(* IEC 61131-3 sources: daoli-st-library/DL_Process (part 3) *)

(* ---- FB_DL_EnergySavingMode.st ---- *)
(*==============================================================================
 * 组件名称 (Component)  : FB_DL_EnergySavingMode
 * 所属子库 (Sublibrary) : DL_Process
 * 当前版本 (Version)    : 1.0.0
 * 组件分类 (Category)   : 功能块（FUNCTION_BLOCK）· 工艺段 · 整线空闲节能编排
 * 兼容性 (Platform)     : CODESYS 3.5 / TwinCAT 3 / 汇川 InoProShop / Machine Expert；
 *                         仅依赖标准库（TON / R_TRIG / LIMIT），气源压力与温度全部经
 *                         引脚注入，块内不读任何外部量、不做任何模拟量通道绑定
 * 功能描述 (Function)   : 以「空闲确认延时 → 节能态（降压 / 停热 / 伺服休眠）→ 唤醒
 *                         缓冲（压力先恢复再放行）」三段编排节能与生产，输出可解释
 *                         的节能标志与累计时长，杜绝「唤醒即放行」造成的低压启动
 * 与既有件边界 (Scope)  : 多台设备轮值由轮值调度件承担；单机运行时长由运行计时件承
 *                         担；本件管整线状态级的能量模式切换与放行门控，不替代任何
 *                         单机控制块，也不下发任何设备级启停指令（只给节能请求位）
 * 状态机规模 (States)   : 四工作态加故障（eRun 0 / eIdleCount 10 / eEco 20 / eWake 30
 *                         / eFault 99）；编号留 10 间隔便于插态
 * 关键算法 (Algorithm)  :
 *   ① 空闲确认：空闲判据须在确认延时内持续为真，中途掉沿立即回运行态并清计时
 *   ② 节能编排：进入顺序固定为「先降压 → 再停热 → 最后伺服休眠」，每步间隔一个台
 *      阶（默认 500 毫秒）；原因是伺服休眠时若气源仍为工作压力，抱闸释放瞬间会顶件
 *   ③ 退出反序：唤醒时严格反序撤销（先撤休眠 → 再撤停热 → 最后恢复压力），保证伺服
 *      再上电时气源已在工作压力附近，不会出现带压顶缸
 *   ④ 唤醒门控：放行须同时满足「压力达节能目标加压裕量」「压力低位请求已撤」「唤醒
 *      缓冲时间走完」三条，防压力表冲高瞬放行
 *   ⑤ 三出口全部为状态派生式，无锁存：既避免单拍标志跨拍残留，也保证任何异常路径
 *      （故障、使能撤销）都会在下一拍自然复位，不需要额外的撤除分支
 *   ⑥ 反馈失效：节能或唤醒期间压力读数触零或非有限值，说明无反馈可用，此时无法确认
 *      压力已恢复，一律禁止放行并锁故障
 * 码位表 (Error codes)  :
 *   16#0005_01C4【信息级】延时或压力参数越界已钳位，不置故障位
 *   16#0005_02F0【故障级】唤醒超时（超过两倍唤醒缓冲仍未达压）
 *   16#0005_02F1【故障级】气源压力反馈缺失（读数为零或非有限值）
 *   16#0005_02F2【故障级】非法状态兜底
 * R32 写入点次序审计 :
 *   bAirPressureLow / bHeatStandby / bServoSleep : 仅在段 9 按状态单点派生（每拍先清零
 *       再按所在阶段置位），状态机内不写，因此不存在同拍多分支写同一量的可能
 *   bReadyToRun : 仅段 9 单点派生（运行态恒真；唤醒态须门控通过）
 *   _uErrorIdInt: ① 首扫清（段 4）→ ② 参数越界（段 2 只进信息码，不写故障码）→ ③ 反馈
 *       缺失（段 6）→ ④ 唤醒超时（段 6）→ ⑤ 非法状态（ELSE）→ ⑥ 复位清（eFault）
 *   _eState     : 每拍只在 CASE 分支出口单点写入；CASE 之外仅段 6 两处监视与段 7 使能
 *       撤销，均在 CASE 之前，次序固定
 *   _tEcoDur    : ① 节能转出拍快照（eEco）→ ② 统计消费拍读取（eWake）→ ③ 复位清
 * 单拍纪律说明 (R24/R25) : 本件节能出口全部为状态派生式（每拍重算、不锁存），因此不
 *       存在单拍标志跨拍残留；唯一具单拍性质的事件是「模式切换」，由切换计数器在节能
 *       转出拍唯一加一承担，不存在预清零与转出拍冲突的问题
 * 验收向量 (Acceptance) :
 *   V1 进入节能：空闲持续达确认延时 → 节能生效为真，同一拍降压请求为真
 *   V2 唤醒门控：节能目标 4.0 巴、裕量 0.2 巴，实测 4.1 巴 → 放行为假（未达 4.2 巴）
 *   V3 唤醒完成：实测 4.25 巴且缓冲走完 → 放行为真，下一拍回运行态
 *   V4 反馈缺失：实测 0.0 巴且节能生效 → 码 02F1、故障态
 *   V5 统计：一次节能持续 300 秒 → 累计节能时长增加 300 秒、切换次数加一
 * 开源溯源 (Origin)     : 参考批控与轻工产线公开手册的能量状态分层与停机分级语义组织，
 *                         只借状态分类与参数域；状态机、反序编排、门控判据、码位与引
 *                         脚契约为本库独立设计，clean-room 不构成衍生作品
 * 红线自检 (Redline)    : R1 零全局表与外部变量引用、零物理地址记号 ✓｜R2 零占位符 ✓
 *                         R3 纯 IEC 61131-3 加标准库 ✓｜R4 非有限值防御、比较全带容差、
 *                         无除法 ✓｜R5 声明行中英双语同行注释 ✓｜R6 五成员逐一有 CASE
 *                         标签且含 ELSE 兜底 ✓｜R7 两沿检测与三定时器全部在 CASE 之外
 *                         无条件刷新 ✓
 * 现场投用须知 (Notes)  :
 *   ① 节能目标压力必须低于工作压力且高于夹具最低夹持压力，低于夹持压力会导致待机
 *      期间工件松脱；建议先按气动原理图核算最低夹持压力再定目标值
 *   ② 唤醒裕量不宜小于压力传感器的重复精度，否则门控会在阈值上下反复抖动；现场
 *      经验值是取传感器精度的三到五倍
 *   ③ 伺服休眠许可由工艺侧给出，本块不判断伺服是否已停稳；若需停机确认，请把停稳
 *      反馈串进许可位，不要在块内加延时猜测
 *   ④ 唤醒缓冲只保证「压力恢复后才放行」，不保证「工件已就位」；来料检测与就位确
 *      认仍由上游工站负责，本块不越权
 * 修订历史 (Revision)   :
 *   2026-11-15  v1.0.0  首版入库（Round 11 · C 泳道 · 工站四件套之四）
 *============================================================================*)

(*------------------------------------------------------------------------------
 * 枚举: E_DL_EcoModeState（归属 FB_DL_EnergySavingMode，同文件发布）
 *   四工作态加故障，每个成员在主状态机中均有同名 CASE 标签（R31 完备性）
 *-----------------------------------------------------------------------------*)
TYPE E_DL_EcoModeState :
(
    eRun       := 0,    // 运行：产线生产，节能出口全撤 / Running, all eco outlets withdrawn
    eIdleCount := 10,   // 空闲确认：等空闲判据持续成立达延时 / Idle confirmation, waiting for the delay
    eEco       := 20,   // 节能：降压、停热、伺服休眠按序投入 / Eco, staged withdrawal of energy
    eWake      := 30,   // 唤醒：按反序恢复并等压力回到工作值 / Wake, reverse restore and pressure gate
    eFault     := 99    // 故障锁存：仅复位沿可退 / Fault latched, only a reset edge leaves
);
END_TYPE

(*------------------------------------------------------------------------------
 * 结构体: ST_DL_EcoStat（归属 FB_DL_EnergySavingMode）
 *   跨周期统计，由调用方持有，本块只累加，掉电保持由上层负责
 *-----------------------------------------------------------------------------*)
TYPE ST_DL_EcoStat :
STRUCT
    tTotalEco    : TIME;                    // 累计节能时长 [毫秒] [Accumulated eco time]
    nSwitchCount : UDINT;                   // 累计模式切换次数 [次] [Mode switch counter]
    tLastEco     : TIME;                    // 上一轮节能时长 [毫秒] [Last eco duration]
END_STRUCT
END_TYPE

FUNCTION_BLOCK FB_DL_EnergySavingMode
VAR_INPUT
    bEnable            : BOOL;              // 使能，FALSE 立即回运行态并撤节能请求 [Enable, FALSE returns to run]
    bReset             : BOOL;              // 复位故障，上升沿受理 [Reset fault on rising edge]
    bLineIdle          : BOOL;              // 产线空闲判据（无料且无作业）[-] [Line idle criterion]
    bWakeRequest       : BOOL;              // 唤醒请求（来料 / 操作员 / 上位机）[-] [Wake-up request]
    fAirPressureAct    : REAL;              // 实际气源压力 [巴]，量程 0.0~10.0 [Actual air pressure, bar]
    fAirPressureEco    : REAL := 4.0;       // 节能目标压力 [巴]，域 0.0~10.0 [Eco target pressure, bar]
    fWakeMargin        : REAL := 0.2;       // 唤醒压力裕量 [巴]，须达目标加裕量 [Wake margin, bar]
    tIdleDelay         : TIME := T#120S;    // 空闲确认延时 [毫秒]，0 表示立即节能 [Idle confirm delay]
    tWakeRamp          : TIME := T#3S;      // 唤醒缓冲（压力恢复等待上限）[毫秒] [Wake ramp allowance]
    bServoSleepPermit  : BOOL;              // 允许伺服休眠，工艺侧给出 [-] [Servo sleep permitted by process]
    bHeatStandbyPermit : BOOL;              // 允许加热转保温或关闭 [-] [Heater standby permitted]
END_VAR
VAR_OUTPUT
    bEcoActive         : BOOL;              // 节能模式生效（节能与唤醒期间均为真）[-] [Eco mode engaged]
    bAirPressureLow    : BOOL;              // 请求降压（送气源比例阀）[-] [Request reduced air pressure]
    bHeatStandby       : BOOL;              // 请求加热转保温或关闭 [-] [Request heater standby]
    bServoSleep        : BOOL;              // 请求伺服休眠 [-] [Request servo sleep]
    bReadyToRun        : BOOL;              // 唤醒完成，可放行生产 [-] [Ready to run after wake]
    eState             : E_DL_EcoModeState; // 主状态机当前态 [-] [Current state]
    bError             : BOOL;              // 故障锁存，需复位清除 [Latched fault]
    uErrorId           : UDINT;             // 事件码或故障码，0 表示无 [Event or fault code]
    tIdleElapsed       : TIME;              // 空闲累计已计时长 [毫秒] [Idle elapsed time]
    tEcoElapsed        : TIME;              // 本次节能已持续时长 [毫秒] [Eco elapsed time]
END_VAR
VAR_IN_OUT
    stStat             : ST_DL_EcoStat;     // 跨周期统计，调用方持有 [Persistent statistics]
END_VAR
VAR
    _eState          : E_DL_EcoModeState := E_DL_EcoModeState.eRun;  // 内部状态寄存器，唯一真值源 [Internal state register]
    _bInit           : BOOL := FALSE;       // 首扫标志，初值 FALSE，判据 NOT _bInit [First-scan flag, R19 pattern]
    _bFaultLatch     : BOOL;                // 故障级锁存，仅复位路径清 [Fault latch, reset path only]
    _uErrorIdInt     : UDINT;               // 故障级码寄存 [Fault-level code register]
    _uInfoCode       : UDINT;               // 本拍信息级码，每拍重算 [Transient info code]
    fEcoEff          : REAL;                // 生效节能目标压力 [巴] [Effective eco pressure, bar]
    fMarginEff       : REAL;                // 生效唤醒裕量 [巴] [Effective wake margin, bar]
    fWakeGate        : REAL;                // 唤醒放行压力门限 [巴] [Wake gate pressure, bar]
    tIdleEff         : TIME;                // 生效空闲延时 [毫秒] [Effective idle delay]
    tWakeEff         : TIME;                // 生效唤醒缓冲 [毫秒] [Effective wake ramp]
    tWakeMaxEff      : TIME;                // 唤醒超时上限（缓冲的两倍）[毫秒] [Wake timeout limit]
    _tEcoDur         : TIME;                // 本次节能实际时长快照 [毫秒] [Eco duration snapshot]
    _bPressFinite    : BOOL;                // 压力读数有限 [-] [Pressure reading finite]
    _bPressMissing   : BOOL;                // 压力反馈缺失判据 [-] [Pressure feedback missing]
    _bWakeGateOk     : BOOL;                // 唤醒放行三条件同时成立 [-] [Wake gate satisfied]
    _bReadyLatch     : BOOL;                // 放行锁存：先放行一拍再转运行态 [Permit latched one scan before returning]
    bIdleIn          : BOOL;                // 空闲计时输入条件，先算后调 [Idle timer input]
    bEcoIn           : BOOL;                // 节能计时输入条件，先算后调 [Eco timer input]
    bWakeIn          : BOOL;                // 唤醒计时输入条件，先算后调 [Wake timer input]
    fbTrigReset      : R_TRIG;              // 复位沿检测 [Reset edge detector]
    fbTrigIdle       : R_TRIG;              // 空闲判据上升沿 [Idle rising edge]
    fbTrigWake       : R_TRIG;              // 唤醒请求上升沿 [Wake request rising edge]
    fbTmoIdle        : TON;                 // 空闲确认计时 [Idle confirmation timer]
    fbTmoEco         : TON;                 // 节能计时兼阶段时钟 [Eco timer and stage clock]
    fbTmoWake        : TON;                 // 唤醒缓冲计时兼阶段时钟 [Wake timer and stage clock]
END_VAR
VAR CONSTANT
    DL_FLOAT_EPS     : REAL := 1.0E-6;      // 浮点判等容差 [-] [Float comparison epsilon]
    DL_PRESSURE_MAX  : REAL := 10.0;        // 压力量程上限 [巴] [Pressure upper bound, bar]
    DL_MARGIN_MAX    : REAL := 5.0;         // 裕量域上限 [巴] [Margin upper bound, bar]
    DL_REAL_MAX      : REAL := 3.4E38;      // 单精度有限值判据幅值 [-] [Finite magnitude bound]
    DL_ECO_GAP1      : TIME := T#500MS;     // 节能与唤醒的第一步台阶 [毫秒] [First stage step]
    DL_ECO_GAP2      : TIME := T#1S;        // 节能与唤醒的第二步台阶 [毫秒] [Second stage step]
    DL_WAKE_FACTOR   : DINT := 2;           // 唤醒超时相对缓冲的倍数 [-] [Wake timeout factor]
    DL_TMO_MAX       : TIME := T#600S;      // 延时参数域上限 [毫秒] [Delay upper bound]
    DL_TIME_MAX      : TIME := T#500H;     // 累计时长饱和上限 [毫秒] [Duration saturation limit]
    DL_SWITCH_MAX    : UDINT := 16#FFFF_FFFE; // 切换次数饱和上限 [次] [Switch counter saturation]
    DL_INFO_LIM_CLAMP: UDINT := 16#0005_01C4; // 01C4 延时或压力参数越界已钳位【信息级】 [Info, parameter clamped]
    DL_ERR_WAKE_TMO  : UDINT := 16#0005_02F0; // 02F0 唤醒超时（压力未恢复）【故障级】 [Fault, wake timeout]
    DL_ERR_PRESS     : UDINT := 16#0005_02F1; // 02F1 气源压力反馈缺失【故障级】 [Fault, pressure feedback missing]
    DL_ERR_STATE     : UDINT := 16#0005_02F2; // 02F2 非法状态兜底【故障级】 [Fault, illegal state]
END_VAR

// ==== 段 1｜信息级码预清零（信息码每拍重算，不跨拍残留） / Info code pre-clear, recomputed every scan
_uInfoCode := 16#0000_0000;                 // 信息级码每拍重算 [Info code recomputed]

// ==== 段 2｜参数钳位（压力、裕量、两个延时，先钳位再进逻辑） / Parameter clamping before any logical use
fEcoEff := fAirPressureEco;                 // 节能目标先取引脚值 [Eco pressure from pin]
IF (fEcoEff < 0.0) OR (fEcoEff > DL_PRESSURE_MAX) THEN
    fEcoEff    := LIMIT(0.0, fEcoEff, DL_PRESSURE_MAX);   // 越界钳到量程内 [Clamped into range]
    _uInfoCode := DL_INFO_LIM_CLAMP;        // 01C4 延时或压力参数越界已钳位【信息级】 [Info, parameter clamped]
END_IF

fMarginEff := fWakeMargin;                  // 裕量先取引脚值 [Margin from pin]
IF (fMarginEff < 0.0) OR (fMarginEff > DL_MARGIN_MAX) THEN
    fMarginEff := LIMIT(0.0, fMarginEff, DL_MARGIN_MAX);  // 越界钳到裕量域内 [Clamped into margin range]
    _uInfoCode := DL_INFO_LIM_CLAMP;        // 01C4 延时或压力参数越界已钳位【信息级】 [Info, parameter clamped]
END_IF

fWakeGate := fEcoEff + fMarginEff;          // 放行门限等于目标加裕量 [Gate = target plus margin]

tIdleEff := tIdleDelay;                     // 空闲延时先取引脚值 [Idle delay from pin]
IF tIdleEff > DL_TMO_MAX THEN
    tIdleEff   := DL_TMO_MAX;               // 超上限钳位 [Clamped to upper bound]
    _uInfoCode := DL_INFO_LIM_CLAMP;        // 01C4 延时或压力参数越界已钳位【信息级】 [Info, parameter clamped]
ELSIF tIdleEff < T#0S THEN
    tIdleEff := T#0S;                       // 负值归零即立即节能 [Negative means immediate]
END_IF

tWakeEff := tWakeRamp;                      // 唤醒缓冲先取引脚值 [Wake ramp from pin]
IF tWakeEff > DL_TMO_MAX THEN
    tWakeEff   := DL_TMO_MAX;               // 超上限钳位 [Clamped to upper bound]
    _uInfoCode := DL_INFO_LIM_CLAMP;        // 01C4 延时或压力参数越界已钳位【信息级】 [Info, parameter clamped]
ELSIF tWakeEff < T#0S THEN
    tWakeEff := T#0S;                       // 负值归零 [Negative clamped to zero]
END_IF

tWakeMaxEff := tWakeEff * DL_WAKE_FACTOR;   // 唤醒超时取缓冲的两倍 [Wake timeout = twice the ramp]

// ==== 段 3｜沿与定时器无条件刷新（R7 红线：严禁置于 IF / CASE 分支内） / Unconditional refresh of edges and timers
fbTrigReset(CLK := bReset);                 // 复位沿 [Reset edge]
fbTrigIdle(CLK := bLineIdle);               // 空闲上升沿 [Idle rising edge]
fbTrigWake(CLK := bWakeRequest);            // 唤醒上升沿 [Wake rising edge]

IF (_eState = E_DL_EcoModeState.eIdleCount) AND bLineIdle THEN
    bIdleIn := TRUE;                        // 空闲确认段且判据仍成立才计时 [Count only while idle persists]
ELSE
    bIdleIn := FALSE;                       // 其余段清零 [Cleared otherwise]
END_IF
fbTmoIdle(IN := bIdleIn, PT := tIdleEff);

IF _eState = E_DL_EcoModeState.eEco THEN
    bEcoIn := TRUE;                         // 节能段计时兼阶段时钟 [Eco timer and stage clock]
ELSE
    bEcoIn := FALSE;                        // 其余段清零 [Cleared otherwise]
END_IF
fbTmoEco(IN := bEcoIn, PT := DL_TIME_MAX);

IF _eState = E_DL_EcoModeState.eWake THEN
    bWakeIn := TRUE;                        // 唤醒段计时兼阶段时钟 [Wake timer and stage clock]
ELSE
    bWakeIn := FALSE;                       // 其余段清零 [Cleared otherwise]
END_IF
fbTmoWake(IN := bWakeIn, PT := DL_TIME_MAX);

// ==== 段 4｜首扫初始化（R19 唯一合法范式：初值 FALSE，判据 NOT，同步后置 TRUE） / First-scan initialisation with the canonical R19 pattern
IF NOT _bInit THEN
    _eState        := E_DL_EcoModeState.eRun;   // 状态回运行 [State to run]
    _bFaultLatch   := FALSE;                // 故障锁存清零 [Fault latch cleared]
    _uErrorIdInt   := 16#0000_0000;         // 故障码清零 [Fault code cleared]
    _tEcoDur       := T#0S;                 // 节能时长快照清零 [Eco snapshot cleared]
    _bReadyLatch   := FALSE;                // 放行锁存复位 [Permit latch reset]
    bEcoActive     := FALSE;                // 节能标志复位 [Eco flag reset]
    bAirPressureLow := FALSE;               // 降压请求复位 [Pressure request reset]
    bHeatStandby   := FALSE;                // 停热请求复位 [Heater request reset]
    bServoSleep    := FALSE;                // 休眠请求复位 [Sleep request reset]
    bReadyToRun    := TRUE;                 // 初始视为可运行 [Initially ready to run]
    bError         := FALSE;                // 故障标志清零 [Error cleared]
    uErrorId       := 16#0000_0000;         // 事件码清零 [Error id cleared]
    tIdleElapsed   := T#0S;                 // 空闲计时清零 [Idle elapsed cleared]
    tEcoElapsed    := T#0S;                 // 节能计时清零 [Eco elapsed cleared]
    stStat.tTotalEco    := T#0S;            // 累计节能时长清零 [Total eco cleared]
    stStat.nSwitchCount := 0;               // 切换次数清零 [Switch counter cleared]
    stStat.tLastEco     := T#0S;            // 上轮节能时长清零 [Last eco cleared]
    _bInit := TRUE;                         // 首扫只做一次 [Runs exactly once]
END_IF

// ==== 段 5｜压力反馈有效性（零读数与非有限值同属「无反馈」，一律按缺失处理） / Pressure feedback validity, zero and non-finite treated alike
_bPressFinite := (fAirPressureAct >= (-DL_REAL_MAX)) AND (fAirPressureAct <= DL_REAL_MAX);
IF (NOT _bPressFinite) OR (fAirPressureAct <= DL_FLOAT_EPS) THEN
    _bPressMissing := TRUE;                 // 无可用反馈 [No usable feedback]
ELSE
    _bPressMissing := FALSE;                // 反馈可用 [Feedback usable]
END_IF

// ==== 段 6｜全局监视：反馈缺失优先，其次唤醒超时（两者都在模式切换之外单点判定） / Global monitors: missing feedback first, then wake timeout
IF bEnable AND (NOT _bFaultLatch) AND _bPressMissing
AND ((_eState = E_DL_EcoModeState.eEco) OR (_eState = E_DL_EcoModeState.eWake)) THEN
    _bFaultLatch := TRUE;                   // 无反馈无法确认恢复，禁止放行 [Cannot confirm recovery, fault]
    _uErrorIdInt := DL_ERR_PRESS;           // 02F1 气源压力反馈缺失【故障级】 [Fault, feedback missing]
    _eState      := E_DL_EcoModeState.eFault;
END_IF

_bWakeGateOk := (_eState = E_DL_EcoModeState.eWake)
            AND (NOT _bPressMissing)
            AND (fAirPressureAct >= (fWakeGate + DL_FLOAT_EPS))
            AND (fbTmoWake.ET >= tWakeEff);   // 门控三条件：压力达标、无缺失、缓冲走完 [Three gate conditions]

IF bEnable AND (NOT _bFaultLatch)
AND (_eState = E_DL_EcoModeState.eWake)
AND (tWakeMaxEff > T#0S)
AND (fbTmoWake.ET > tWakeMaxEff)
AND (NOT _bWakeGateOk) THEN
    _bFaultLatch := TRUE;                   // 缓冲两倍仍未达压，锁故障 [Pressure not restored, fault]
    _uErrorIdInt := DL_ERR_WAKE_TMO;        // 02F0 唤醒超时【故障级】 [Fault, wake timeout]
    _eState      := E_DL_EcoModeState.eFault;
END_IF

// ==== 段 7｜使能撤销（FALSE 立即回运行态，节能出口由段 9 自然撤销） / Disable path returns to run, eco outlets drop by derivation
IF NOT bEnable THEN
    _eState := E_DL_EcoModeState.eRun;      // 立即回运行态 [Immediately back to run]
    _tEcoDur := T#0S;                       // 时长快照作废 [Snapshot invalidated]
END_IF

// ==== 段 8｜主状态机（ENUM 加 CASE 加 ELSE 兜底，五成员逐一有标签） / Main state machine, every member has its own label
CASE _eState OF
    E_DL_EcoModeState.eRun: // 运行：等空闲判据上升沿
        IF fbTrigIdle.Q AND bEnable AND (NOT _bFaultLatch) THEN
            _uErrorIdInt := 16#0000_0000;   // 进入确认前无故障 [No fault before confirmation]
            _eState      := E_DL_EcoModeState.eIdleCount;
        END_IF

    E_DL_EcoModeState.eIdleCount: // 空闲确认：判据中途掉沿立即回运行
        IF NOT bLineIdle THEN
            _eState := E_DL_EcoModeState.eRun;     // 判据失守，回运行态 [Idle criterion lost, back to run]
        ELSIF fbTmoIdle.Q THEN
            _tEcoDur := T#0S;               // 新一轮节能，时长快照清零 [New eco round, snapshot cleared]
            _eState  := E_DL_EcoModeState.eEco;
        END_IF

    E_DL_EcoModeState.eEco: // 节能：三段按阶投入，唤醒请求或来料即转唤醒
        IF fbTrigWake.Q OR (NOT bLineIdle) THEN
            _tEcoDur     := fbTmoEco.ET;    // 转出拍快照节能时长（定时器出段即清零）[Snapshot before the timer resets]
            _bReadyLatch := FALSE;          // 新的唤醒过程，放行锁存复位 [Permit latch reset]
            _eState      := E_DL_EcoModeState.eWake;
        END_IF

    E_DL_EcoModeState.eWake: // 唤醒：三条件成立先放行一拍，下一拍才转运行
        IF _bWakeGateOk AND (NOT _bReadyLatch) THEN
            _bReadyLatch := TRUE;           // 本拍放行（bReadyToRun 由出口派生为真）[Permit for this scan only]
        ELSIF _bWakeGateOk AND _bReadyLatch THEN
            IF stStat.nSwitchCount < DL_SWITCH_MAX THEN
                stStat.nSwitchCount := stStat.nSwitchCount + 1;   // 模式切换计数，本拍唯一加一 [Switch counter, single increment]
            END_IF
            stStat.tLastEco := _tEcoDur;    // 上一轮节能时长 [Last eco duration]
            IF stStat.tTotalEco < DL_TIME_MAX THEN
                stStat.tTotalEco := stStat.tTotalEco + _tEcoDur;  // 累计节能时长饱和累加 [Total eco accumulated]
            END_IF
            _bReadyLatch := FALSE;          // 转出即复位 [Reset on exit]
            _eState      := E_DL_EcoModeState.eRun;
        ELSIF NOT _bWakeGateOk THEN
            _bReadyLatch := FALSE;          // 门控失守（压力回落）则撤销放行 [Gate lost, permit revoked]
        END_IF

    E_DL_EcoModeState.eFault: // 故障：等复位沿，复位后清码回运行
        IF fbTrigReset.Q THEN
            _bFaultLatch := FALSE;          // 锁存解除 [Latch released]
            _uErrorIdInt := 16#0000_0000;   // 故障码清零 [Fault code cleared]
            _tEcoDur     := T#0S;           // 时长快照作废 [Snapshot invalidated]
            _bReadyLatch := FALSE;          // 放行锁存复位 [Permit latch reset]
            _eState      := E_DL_EcoModeState.eRun;
        END_IF

    ELSE // 非法枚举值兜底：回安全态并锁故障（节能出口由段 9 派生为假）
        _bFaultLatch := TRUE;               // 兜底锁存 [Fallback latch]
        _uErrorIdInt := DL_ERR_STATE;       // 02F2 非法状态兜底【故障级】 [Fault, illegal state]
        _eState      := E_DL_EcoModeState.eFault;
END_CASE

// ==== 段 9｜出口派生（三个节能出口与放行位全部按状态与阶段单点派生） / Outlets derived from state and stage at a single point
bAirPressureLow := FALSE;                   // 先清零再按阶段置位 [Pre-cleared, then set by stage]
bHeatStandby    := FALSE;
bServoSleep     := FALSE;

IF _eState = E_DL_EcoModeState.eEco THEN
    bAirPressureLow := TRUE;                // 第一步：先降压（伺服仍带电，防带压休眠）[Step 1: reduce pressure first]
    IF (fbTmoEco.ET >= DL_ECO_GAP1) AND bHeatStandbyPermit THEN
        bHeatStandby := TRUE;               // 第二步：降压稳定后再停热 [Step 2: heater standby after pressure settled]
    END_IF
    IF (fbTmoEco.ET >= DL_ECO_GAP2) AND bServoSleepPermit THEN
        bServoSleep := TRUE;                // 第三步：最后才允许伺服休眠 [Step 3: servo sleep last]
    END_IF
ELSIF _eState = E_DL_EcoModeState.eWake THEN
    IF fbTmoWake.ET < DL_ECO_GAP1 THEN
        bHeatStandby   := TRUE;             // 反序第一步：先撤休眠，其余保持不动作 [Reverse step 1: sleep released first]
        bAirPressureLow := TRUE;            // 压力仍处低位 [Pressure still low]
    ELSIF fbTmoWake.ET < DL_ECO_GAP2 THEN
        bAirPressureLow := TRUE;            // 反序第二步：停热已撤，压力仍低位 [Reverse step 2: heater restored, pressure low]
    END_IF
    // 反序第三步：压力请求撤除（三出口全假），由气源比例阀自行回到工作压力
END_IF

bEcoActive  := (_eState = E_DL_EcoModeState.eEco)
            OR (_eState = E_DL_EcoModeState.eWake);   // 节能与唤醒期间均视为节能投入 [Engaged during eco and wake]

bReadyToRun := (_eState = E_DL_EcoModeState.eRun)
            OR _bReadyLatch;                // 运行态恒可运行；唤醒态须放行锁存已置 [Ready in run, or when latched in wake]

IF _eState = E_DL_EcoModeState.eWake THEN
    tEcoElapsed := _tEcoDur;                // 唤醒期间显示本轮节能已持续时长 [Show the finished eco duration]
ELSE
    tEcoElapsed := fbTmoEco.ET;             // 其余时段按节能定时器已历时 [Eco timer elapsed otherwise]
END_IF
tIdleElapsed := fbTmoIdle.ET;               // 空闲确认已计时长 [Idle confirmation elapsed]

eState := _eState;                          // 状态镜像 [State mirror]
bError := _bFaultLatch;                     // 故障级派生式（R21）[Fault-level derived form]
IF _bFaultLatch THEN
    uErrorId := _uErrorIdInt;               // 故障级码优先透出 [Fault code wins]
ELSE
    uErrorId := _uInfoCode;                 // 无故障时透出信息级码 [Info code otherwise]
END_IF

// ==== 段 10｜现场提示（调试与验收要点，不参与逻辑） / Field notes, no logic impact
//   1 三个节能出口均为派生式：任何时刻读到的值都与当前状态严格一致，不存在「已撤
//     状态但出口还挂着」的中间态，这是排查「节能撤不掉」类问题的前提；
//   2 进入节能后第一步只降压，停热与休眠各隔一个台阶（默认 500 毫秒），台阶时长
//     由常量给定，若现场气源响应慢，改常量而不是在逻辑里加延时；
//   3 唤醒超时取缓冲的两倍：一倍用于压力恢复，另一倍留给比例阀回差与管路充气，
//     超过两倍仍未达压说明气源或阀件有问题，此时锁故障比继续等待更有价值；
//   4 切换次数在节能转出拍加一，与累计时长同一拍结算，两者可在上位机互校。
END_FUNCTION_BLOCK

(* ---- FB_DL_FrameSealDispenseSeq.st ---- *)
(*==============================================================================
 * 组件名称 (Component)  : FB_DL_FrameSealDispenseSeq
 * 所属子库 (Sublibrary) : DL_Process
 * 当前版本 (Version)    : 1.0.0
 * 兼容性   (Platform)   : CODESYS 3.5+ / TwinCAT 3 / 汇川 InoProShop / 施耐德 Machine Expert
 *                         仅依赖 Standard.library（TON / R_TRIG / ABS），零厂商私有库
 * 功能描述 (Function)   : 装框打胶顺控：eIdle → eHome（打胶头回参考）→ ePurge（预挤胶，废胶接料）
 *                         → eDispense（分段打胶，按 nSegCount 段推进，每段校核胶量）→ ePress
 *                         （压合到位）→ eCure（固化窗计时）→ eDone。断胶检测：eDispense 中
 *                         bGlueFlow 连续 tFlowGapMax 无信号 → 判断胶故障并**立即停止打胶并锁存**
 *                         （安全侧：断胶继续走会做出废件且可能把胶漏到设备上）。
 * 取舍声明 (Trade-off)  : **单段胶量超差不中断打胶**：某段胶量偏差超 fDoseTolPct 时该段计 NG，
 *                         但**继续打完剩余段**——半截停止会让整框报废，而打完剩下段至少能拿到
 *                         完整胶道供返修与工艺分析；NG 结论在循环结束时以 nNgSegCount 与 eCause
 *                         = eDoseNg 一并给出。这一取舍与「断胶立即停」并不矛盾：胶量超差是
 *                         **质量降级**，断胶是**工艺不可继续**，前者可回收后者不可。
 * 接口     (Interface)  : 输入 bStart 启动电平、bHomeDone 回参到位、bPurgeDone、bSegDone 段完成沿、
 *                         bPressDone 压合到位、bGlueFlow 胶流在位、fGlueDoseG 段实测胶量、
 *                         fDoseTgtG 段目标胶量、fDoseTolPct 胶量容差百分比、nSegCount 段数、
 *                         六个时间量（回参/预挤/断胶/压合/固化及其超时）、bReset 复位；
 *                         输出 eState、eCause、bGlueOn 打胶阀命令、bPressCmd 压合命令、bPurgeCmd、
 *                         bHomeCmd、nSegDone 已完成段数、nNgSegCount NG 段累计（锁存量，复位不清零）、
 *                         bBatchNg 本批次 NG 结论、bCycleDone、bError、nErrId。
 * 边界     (Boundary)   : ① 组态闸：fDoseTolPct <= 0.0、fDoseTgtG <= 0.0、nSegCount = 0、任一时长
 *                         <= T#0S、时长配比越界（超时 <= 工艺时长）或任一浮点引脚 NaN → 故障锁存；
 *                         ② TON 五枚 + R_TRIG 三枚段 0 无条件刷新，IN 均由相位派生（R228A）；
 *                         ③ **NG 计数为锁存量，复位不清零**（批次台账语义）；窗内极值类当拍量才清；
 *                         ④ 断胶判据只在 eDispense 相内使能，离开该相自动复位（R228B）；
 *                         ⑤ 故障相迁出唯一路径 = bReset 上升沿；⑥ 零全局耦合（无 GVL / 无物理地址）。
 * 定时器清单 (Timers)   : 本件 5 枚 TON + 3 枚 R_TRIG（较派单 4+2 各多一枚，理由：tonFlow 的 IN
 *                         必须随 bGlueFlow 在相内独立复位，不能与相计时合并；段完成沿 bSegDone
 *                         必须独立成沿实例，不能与启动沿或复位沿合并），全部段 0 无条件调用。
 * 解除式   (Release)    : bReset 上升沿 ∧ 组态合法 ∧ 无断胶（bGlueFlow 当拍为真，R240 范式）。
 *                         自证可满足（终审两式 1）：五枚 TON 的 IN 挂相位，故障相内恒假 → Q 恒假；
 *                         恢复供胶后 bGlueFlow 为真即达，无恒假因子。
 * 码表     (Codes)      : 16#0005_03A7 故障级：装框打胶顺控故障总码（组态非法 / 回参超时 / 预挤超时 /
 *                         断胶 / 压合超时 / 固化超时 / 非法相位），锁存至 bReset 上升沿，归因由
 *                         eCause 承载（R190 单件单总码）；16#0005_04CF 信息级：批次正常完成。
 *                         归因说明：eCause 亦承载**非故障**的批次质量归因 eDoseNg（胶量超差但循环
 *                         走完），此时 bError 恒为 FALSE——HMI 必须用 bError 判故障、用 eCause 判
 *                         质量归因，不得以 eCause 非零视为故障（R191 名实双出口）。
 *                         加码反证（R90）：批次完成时 bCycleDone 由相位派生，「完成态驻留」与之同值；
 *                         且 NG 结论 bBatchNg 也会在完成态保持，出口组合无法区分「刚完成一次」
 *                         与「长期驻留完成态」，故立一码记录每次完成沿。
 *                         码段说明：0005 段故障子带 03xx / 信息子带 04xx，本件取 03A7 / 04CF
 *                         （源码实扫该两槽为空，续接同子带已用最大值，未回填碎片孔洞）。
 * 开源溯源 (Origin)     : 道莅自研 clean-room（参考光伏组件装框打胶工艺与公开参数域，
 *                         零代码行复制；自研行业池）
 * 修订历史 (Revision)   : 2026-11-19  v1.0.0  R45 首版（批次 4 · 序号 19）
 *==============================================================================*)

TYPE E_DL_FsdState :
(
    eIdle     := 0,     // 待启动 / Idle, awaiting start
    eHome     := 10,    // 打胶头回参考 / Dispenser homing
    ePurge    := 20,    // 预挤胶（废胶接料） / Purging to the waste cup
    eDispense := 30,    // 分段打胶 / Segmented dispensing
    ePress    := 40,    // 压合 / Pressing
    eCure     := 50,    // 固化窗计时 / Curing window
    eDone     := 60,    // 批次完成 / Batch done
    eFault    := 90     // 故障锁存相 / Fault latched phase
);
END_TYPE

TYPE E_DL_FsdCause :
(
    eNone       := 0,   // 无故障成因 / No cause
    eCfgIllegal := 1,   // 组态非法 / Illegal configuration
    eHomeTmo    := 2,   // 回参超时 / Homing timeout
    ePurgeTmo   := 3,   // 预挤超时 / Purge timeout
    eNoGlue     := 4,   // 断胶（流量信号消失超时） / Glue flow lost
    ePressTmo   := 5,   // 压合超时 / Press timeout
    eCureTmo    := 6,   // 固化超时 / Cure timeout
    eDoseNg     := 7,   // 胶量超差（非故障，批次质量归因） / Dose out of tolerance, quality attribution only
    ePhaseBad   := 8    // 非法相位兜底 / Illegal phase fallback
);
END_TYPE

FUNCTION_BLOCK FB_DL_FrameSealDispenseSeq
VAR_INPUT
    bStart        : BOOL := FALSE;        // 启动电平（落沿等于撤启动） [-] / Start level, falling edge means abort
    bHomeDone     : BOOL := FALSE;        // 打胶头回参考到位 [-] / Dispenser homed
    bPurgeDone    : BOOL := FALSE;        // 预挤完成 [-] / Purge finished
    bSegDone      : BOOL := FALSE;        // 当前段完成，上升沿受理一段 [-] / Segment done, rising edge accepts one segment
    bPressDone    : BOOL := FALSE;        // 压合到位 [-] / Pressed in position
    bGlueFlow     : BOOL := FALSE;        // 胶流在位（断胶判据） [-] / Glue flow present
    fGlueDoseG    : REAL := 0.0;          // 当前段累计胶量 [g] / Accumulated dose of the current segment [g]
    fDoseTgtG     : REAL := 5.0;          // 段目标胶量，域 > 0.0 [g] / Segment target dose, domain > 0.0 [g]
    fDoseTolPct   : REAL := 5.0;          // 段胶量容差百分比，域 > 0.0 [%] / Segment dose tolerance, domain > 0.0 [%]
    nSegCount     : INT := 8;             // 段数（正整数），域 > 0 [段] / Segment count, domain > 0 [seg]
    tHomeMax      : TIME := T#20S;        // 回参超时，域 > T#0S [ms] / Homing timeout [ms]
    tPurge        : TIME := T#3S;         // 预挤工艺时长，域 > T#0S [ms] / Purge process time [ms]
    tPurgeMax     : TIME := T#8S;         // 预挤超时，域 > tPurge [ms] / Purge timeout [ms]
    tFlowGapMax   : TIME := T#300MS;      // 断胶判定时长（无胶流超时），域 > T#0S [ms] / Glue-flow gap limit [ms]
    tPressMax     : TIME := T#15S;        // 压合超时，域 > T#0S [ms] / Press timeout [ms]
    tCure         : TIME := T#30S;        // 固化工艺时长，域 > T#0S [ms] / Cure process time [ms]
    tCureMax      : TIME := T#60S;        // 固化超时，域 > tCure [ms] / Cure timeout [ms]
    bReset        : BOOL := FALSE;        // 复位命令，上升沿清故障（不清 NG 台账） [-] / Reset clears fault, not the NG ledger
END_VAR
VAR_OUTPUT
    eState        : E_DL_FsdState;        // 状态出口，段 6 单点映射 / State outlet
    eCause        : E_DL_FsdCause;        // 成因出口（故障归因或批次质量归因） / Cause outlet, fault or quality attribution
    bGlueOn       : BOOL;                 // 打胶阀命令（仅 eDispense 相） [-] / Glue valve command, dispense phase only
    bPressCmd     : BOOL;                 // 压合命令（仅 ePress 相） [-] / Press command, press phase only
    bPurgeCmd     : BOOL;                 // 预挤命令（仅 ePurge 相） [-] / Purge command, purge phase only
    bHomeCmd      : BOOL;                 // 回参命令（仅 eHome 相） [-] / Homing command, home phase only
    nSegDone      : INT;                  // 已完成段数 [段] / Segments completed [seg]
    nNgSegCount   : INT;                  // NG 段累计（锁存量，复位不清零） [段] / NG segment total, latched, kept across resets
    bBatchNg      : BOOL;                 // 本批次 NG 结论（NG 段 > 0） [-] / Batch NG verdict
    bCycleDone    : BOOL;                 // 批次完成标志 [-] / Batch done flag
    bError        : BOOL;                 // 故障锁存标志 [-] / Fault latch flag
    nErrId        : UDINT;                // 事件码，0 = 无事件 / Event code, 0 = no event
END_VAR
VAR
    _eState       : E_DL_FsdState := E_DL_FsdState.eIdle;   // 内部相位（CASE 唯一写入目标） / Internal phase
    _eCause       : E_DL_FsdCause := E_DL_FsdCause.eNone;   // 成因锁存（锁存量） / Latched cause
    tonHome       : TON;                  // 回参计时（PT = 超时），段 0 无条件调用 / Homing timer
    tonPurge      : TON;                  // 预挤计时（PT = 超时），段 0 无条件调用 / Purge timer
    tonFlow       : TON;                  // 断胶计时（IN 随胶流独立复位），段 0 无条件调用 / Glue-gap timer
    tonPress      : TON;                  // 压合计时（PT = 超时），段 0 无条件调用 / Press timer
    tonCure       : TON;                  // 固化计时（PT = 超时），段 0 无条件调用 / Cure timer
    rtSeg         : R_TRIG;               // 段完成沿实例，段 0 无条件调用 / Segment-done edge
    rtStart       : R_TRIG;               // 启动沿实例，段 0 无条件调用 / Start edge
    rtReset       : R_TRIG;               // 复位沿实例，段 0 无条件调用 / Reset edge
    _nSegDone     : INT;                  // 已完成段计数（锁存量） [段] / Completed segment counter, latched
    _nNgSeg       : INT;                  // NG 段计数（锁存量，复位不清零） [段] / NG segment counter, kept across resets
    _fDoseDevPct  : REAL;                 // 段胶量相对偏差当拍量 [%] / Segment relative dose deviation [%]
    _bNonFin      : BOOL;                 // 输入非有限当拍量 [-] / Non-finite input this scan
    _bCfgBad      : BOOL;                 // 组态非法当拍量 [-] / Illegal configuration
    _bFault       : BOOL;                 // 故障锁存位（锁存量） / Latched fault bit
    _uFault       : UDINT;                // 故障码锁存（锁存量） / Latched fault code
    _uInfo        : UDINT;                // 信息码，每拍重算 / Info code, recomputed each scan
END_VAR
VAR CONSTANT
    DL_FLOAT_EPS : REAL := 1.0E-6;        // 浮点判零容差（除子统一口径） [无量纲] / Float epsilon for zero tests
    DL_PCT_SCALE : REAL := 100.0;         // 百分比换算常数 [%] / Percentage scaling constant [%]
END_VAR

(* —— 段 0：当拍判据派生 + 5 枚 TON 与 3 枚 R_TRIG 无条件周期刷新 —— *)
_bNonFin := (fGlueDoseG <> fGlueDoseG) OR (fDoseTgtG <> fDoseTgtG) OR (fDoseTolPct <> fDoseTolPct);   // NaN 自反判（判等禁令唯一例外） / NaN self-reflexive tests
IF fDoseTgtG > DL_FLOAT_EPS THEN                                                                       // 除零前置判 / Divide-by-zero guard
    _fDoseDevPct := (ABS(fGlueDoseG - fDoseTgtG) / fDoseTgtG) * DL_PCT_SCALE;                          // 段胶量相对偏差 / Segment relative dose deviation
ELSE
    _fDoseDevPct := DL_PCT_SCALE;                                                                       // 目标退化按最差偏差处理（组态闸已拦） / Degenerate target treated as worst deviation
END_IF
_bCfgBad := (fDoseTolPct <= 0.0) OR (fDoseTgtG <= 0.0) OR (nSegCount <= 0)                              // 容差与段数组态闸（R151） / Tolerance and segment-count gates
            OR (tHomeMax <= T#0S) OR (tPurge <= T#0S) OR (tPurgeMax <= tPurge)                          // 回参与预挤时间闸 / Homing and purge gates
            OR (tFlowGapMax <= T#0S) OR (tPressMax <= T#0S)                                             // 断胶与压合时间闸 / Glue-gap and press gates
            OR (tCure <= T#0S) OR (tCureMax <= tCure);                                                  // 固化时间配比闸 / Cure time gates
rtSeg(CLK := bSegDone);                                                                                 // 段完成沿，每拍必调（R228A） / Segment edge
rtStart(CLK := bStart);                                                                                 // 启动沿，每拍必调 / Start edge
rtReset(CLK := bReset);                                                                                 // 复位沿，每拍必调 / Reset edge
tonHome(IN := (_eState = E_DL_FsdState.eHome), PT := tHomeMax);                                          // 回参计时（IN 绑相位） / Homing timer
tonPurge(IN := (_eState = E_DL_FsdState.ePurge), PT := tPurgeMax);                                       // 预挤计时（IN 绑相位） / Purge timer
tonFlow(IN := (_eState = E_DL_FsdState.eDispense) AND (NOT bGlueFlow), PT := tFlowGapMax);                // 断胶计时（相内随胶流复位） / Glue-gap timer
tonPress(IN := (_eState = E_DL_FsdState.ePress), PT := tPressMax);                                       // 压合计时（IN 绑相位） / Press timer
tonCure(IN := (_eState = E_DL_FsdState.eCure), PT := tCureMax);                                          // 固化计时（IN 绑相位） / Cure timer

(* —— 段 1：单拍量预清零（锁存量不入清单，R107） —— *)
_uInfo     := 16#0000_0000;        // 信息码每拍重算 / Info recomputed every scan
nSegDone   := _nSegDone;           // 完成段数镜像（锁存量回放） / Segment-done mirror
nNgSegCount := _nNgSeg;            // NG 台账镜像（锁存量回放，复位不清零） / NG ledger mirror
bBatchNg   := (_nNgSeg > 0);       // 批次 NG 结论由台账派生（名实同源） / Batch verdict derived from the ledger
nErrId     := 16#0000_0000;        // 事件码缺省无事件 / Event code default none
bError     := FALSE;               // 故障标志每拍预清，故障分支同拍置位（R45 配对） / Flag preset

(* —— 段 2：复位沿 + 组态域闸 + 非有限闸 —— *)
IF rtReset.Q THEN                                                        // 当拍复位沿 / current-scan reset edge
    _bFault := FALSE;                                                    // 清故障锁存位（锁存量） / Clear fault latch
    _uFault := 16#0000_0000;                                             // 清故障锁存码（锁存量） / Clear latched code
    _eCause := E_DL_FsdCause.eNone;                                      // 清成因（锁存量） / Clear latched cause
    IF _eState = E_DL_FsdState.eFault THEN
        _eState := E_DL_FsdState.eIdle;                                  // 故障相迁出唯一路径 / Sole exit from fault phase
    END_IF
END_IF
IF _bCfgBad THEN                                                         // 组态域闸 / Configuration gate
    _uFault := 16#0005_03A7;                                             // 故障级：装框打胶顺控故障总码 / Fault-level: dispensing sequence fault code
    _bFault := TRUE;
    bError  := TRUE;                                                     // 故障标志同拍置位（R45 配对） / Error flag set same scan
    _eCause := E_DL_FsdCause.eCfgIllegal;                                // 归因：组态非法 / Cause: illegal configuration
END_IF
IF (NOT _bFault) AND _bNonFin THEN                                       // 输入非有限 / Non-finite input
    _uFault := 16#0005_03A7;
    _bFault := TRUE;
    bError  := TRUE;
    _eCause := E_DL_FsdCause.eCfgIllegal;                                // 归因：组态非法（含非有限输入） / Cause: illegal configuration with non-finite input
END_IF
IF (NOT _bFault) AND tonFlow.Q THEN                                      // 断胶：立即停止打胶并锁存（安全侧） / Glue lost, stop immediately and latch
    _uFault := 16#0005_03A7;
    _bFault := TRUE;
    bError  := TRUE;
    _eCause := E_DL_FsdCause.eNoGlue;                                    // 归因：断胶 / Cause: glue flow lost
END_IF

(* —— 段 3：相超时判据（各成因独立赋值点，R190） —— *)
IF (NOT _bFault) AND tonHome.Q THEN
    _uFault := 16#0005_03A7;
    _bFault := TRUE;
    bError  := TRUE;
    _eCause := E_DL_FsdCause.eHomeTmo;                                   // 归因：回参超时 / Cause: homing timeout
END_IF
IF (NOT _bFault) AND tonPurge.Q THEN
    _uFault := 16#0005_03A7;
    _bFault := TRUE;
    bError  := TRUE;
    _eCause := E_DL_FsdCause.ePurgeTmo;                                  // 归因：预挤超时 / Cause: purge timeout
END_IF
IF (NOT _bFault) AND tonPress.Q THEN
    _uFault := 16#0005_03A7;
    _bFault := TRUE;
    bError  := TRUE;
    _eCause := E_DL_FsdCause.ePressTmo;                                  // 归因：压合超时 / Cause: press timeout
END_IF
IF (NOT _bFault) AND tonCure.Q THEN
    _uFault := 16#0005_03A7;
    _bFault := TRUE;
    bError  := TRUE;
    _eCause := E_DL_FsdCause.eCureTmo;                                   // 归因：固化超时 / Cause: cure timeout
END_IF

(* —— 段 4：段级胶量校核（NG 只记台账不中断，头注释取舍声明） —— *)
IF (NOT _bFault) AND (_eState = E_DL_FsdState.eDispense) AND rtSeg.Q THEN
    IF _nSegDone < nSegCount THEN                                        // 段数未满才受理 / Accept only while segments remain
        _nSegDone := _nSegDone + 1;                                      // 累计完成段 / Count the segment
        IF _fDoseDevPct > fDoseTolPct THEN                               // 胶量超差：记 NG 但继续打（不中断） / Over tolerance, record NG and continue
            IF _nNgSeg < 32767 THEN
                _nNgSeg := _nNgSeg + 1;                                  // NG 台账递增（锁存量） / NG ledger increment, latched
            END_IF
            _eCause := E_DL_FsdCause.eDoseNg;                            // 质量归因（非故障，bError 保持 FALSE） / Quality attribution, not a fault
        END_IF
    END_IF
END_IF

(* —— 段 5：故障解除式（R240 全当拍量；NG 台账不受复位影响） —— *)
IF rtReset.Q AND (NOT _bCfgBad) AND (NOT _bNonFin) AND bGlueFlow THEN
    _bFault := FALSE;                                                    // 清故障锁存位（锁存量） / Clear fault latch
    _uFault := 16#0000_0000;                                             // 清故障锁存码（锁存量） / Clear latched code
    _eCause := E_DL_FsdCause.eNone;                                      // 清成因（锁存量，NG 台账仍保留） / Clear cause, NG ledger preserved
END_IF

(* —— 段 5A：故障锁存相位迁移闸 —— *)
IF _bFault AND (_eState <> E_DL_FsdState.eFault) THEN
    _eState := E_DL_FsdState.eFault;                                     // 锁存即入故障相 / Latch enters fault phase
END_IF

(* —— 段 6：相位机（ENUM 全成员显式标签 + ELSE 兜底，R128） —— *)
CASE _eState OF

E_DL_FsdState.eIdle:
    IF rtStart.Q AND (NOT _bFault) THEN                                  // 出口 1：启动沿 / Start edge
        _nSegDone := 0;                                                  // 新批次清完成段（台账 nNgSeg 不清） / Reset segment progress, NG ledger kept
        _eState := E_DL_FsdState.eHome;
    ELSIF _bFault THEN                                                   // 出口 2：故障锁存 / Fault latched
        _eState := E_DL_FsdState.eFault;
    END_IF

E_DL_FsdState.eHome:
    IF bHomeDone THEN                                                    // 出口 1：回参到位 / Homed
        _eState := E_DL_FsdState.ePurge;
    ELSIF NOT bStart THEN                                                // 出口 2：撤启动（前置消失，R98） / Start released
        _eState := E_DL_FsdState.eIdle;
    END_IF

E_DL_FsdState.ePurge:
    IF (bPurgeDone OR (tonPurge.ET >= tPurge)) THEN                      // 出口 1：预挤完成或工艺时长届满 / Purge done or process time reached
        _eState := E_DL_FsdState.eDispense;
    ELSIF NOT bStart THEN                                                // 出口 2：撤启动 / Start released
        _eState := E_DL_FsdState.eIdle;
    END_IF

E_DL_FsdState.eDispense:
    IF _nSegDone >= nSegCount THEN                                       // 出口 1：全部段完成 / All segments done
        _eState := E_DL_FsdState.ePress;
    ELSIF NOT bStart THEN                                                // 出口 2：撤启动 / Start released
        _eState := E_DL_FsdState.eIdle;
    END_IF

E_DL_FsdState.ePress:
    IF bPressDone THEN                                                   // 出口 1：压合到位 / Pressed in position
        _eState := E_DL_FsdState.eCure;
    ELSIF NOT bStart THEN                                                // 出口 2：撤启动 / Start released
        _eState := E_DL_FsdState.eIdle;
    END_IF

E_DL_FsdState.eCure:
    IF tonCure.ET >= tCure THEN                                          // 出口 1：固化时长届满 / Cure time reached
        _uInfo := 16#0005_04CF;                                          // 信息级：批次正常完成 / Info: batch completed
        _eState := E_DL_FsdState.eDone;
    ELSIF NOT bStart THEN                                                // 出口 2：撤启动 / Start released
        _eState := E_DL_FsdState.eIdle;
    END_IF

E_DL_FsdState.eDone:
    bCycleDone := TRUE;                                                  // 完成相保持完成标志 / Hold done flag in done phase
    IF NOT bStart THEN                                                   // 出口 1：撤启动回空闲 / Start released returns idle
        _eState := E_DL_FsdState.eIdle;
    ELSIF _bFault THEN                                                   // 出口 2：故障锁存 / Fault latched
        _eState := E_DL_FsdState.eFault;
    END_IF

E_DL_FsdState.eFault:
    ;                                                                     // 故障相：仅段 5 复位沿可迁出 / Only the reset edge leaves this phase

ELSE
    _uFault := 16#0005_03A7;                                             // 故障级：非法相位兜底（归并总码） / Illegal-phase fallback
    _bFault := TRUE;
    bError  := TRUE;
    _eCause := E_DL_FsdCause.ePhaseBad;                                  // 归因：非法相位 / Cause: illegal phase
    _eState := E_DL_FsdState.eFault;

END_CASE

(* —— 段 7：出口单点映射（名实同源；锁存码回放；故障相命令全落） —— *)
IF _bFault THEN
    bGlueOn    := FALSE;                                                 // 故障相：打胶阀关（断胶/超时均不得继续打胶） / Glue valve closed in fault
    bPressCmd  := FALSE;                                                 // 故障相：压合命令撤 / Press command released in fault
    bPurgeCmd  := FALSE;                                                 // 故障相：预挤命令撤 / Purge command released in fault
    bHomeCmd   := FALSE;                                                 // 故障相：回参命令撤 / Home command released in fault
    bCycleDone := FALSE;                                                 // 故障相不宣称完成 / No completion claim in fault
ELSE
    bGlueOn    := (_eState = E_DL_FsdState.eDispense);                   // 打胶阀仅打胶相开 / Glue valve only while dispensing
    bPressCmd  := (_eState = E_DL_FsdState.ePress);                      // 压合仅压合相 / Press only in press phase
    bPurgeCmd  := (_eState = E_DL_FsdState.ePurge);                      // 预挤仅预挤相 / Purge only in purge phase
    bHomeCmd   := (_eState = E_DL_FsdState.eHome);                       // 回参仅回参相 / Home only in home phase
END_IF
IF _bFault THEN
    nErrId := _uFault;                                                   // 故障锁存码回放 / Replay latched fault code
ELSE
    nErrId := _uInfo;                                                    // 信息码 / Info code
END_IF
bError := _bFault;                                                       // 故障标志与锁存同源（名实双出口，R191） / Flag from latch
eState := _eState;                                                       // 状态出口 / State outlet
eCause := _eCause;                                                       // 成因出口 / Cause outlet

END_FUNCTION_BLOCK

(* ---- FB_DL_LaminatorZoneSync.st ---- *)
(*==============================================================================
 * 组件名称 (Component)  : FB_DL_LaminatorZoneSync
 * 所属子库 (Sublibrary) : DL_Process
 * 当前版本 (Version)    : 1.0.0
 * 兼容性   (Platform)   : CODESYS 3.5+ / TwinCAT 3 / 汇川 InoProShop / 施耐德 Machine Expert
 *                         仅依赖 Standard.library（TON / R_TRIG），零厂商私有库
 * 功能描述 (Function)   : 层压机多温区联动升温。
 *                         把 1..4 个温区当作一个**联动体**（非独立温控）来推：同一设定、统一分级投切、
 *                         统一限温差，避免各区各自为政造成"局部过冲 → 材料应力"。
 *                         三段语义：
 *                           ① **分级投切**：按"设定 − 平均实测"的偏差分三级
 *                              Δ > fDevStage3 → 三级（满功率）；Δ > fDevStage2 → 二级；
 *                              Δ > fDevStage1 → 一级；否则零级（保温/停加热）。
 *                              分级门槛必须单调递减（fDevStage3 > fDevStage2 > fDevStage1 > 0），否则组态非法；
 *                           ② **最小驻留**：每次换级后 tStageMin 内不再换级（防调功器被高频投切打坏）；
 *                           ③ **区间温差联锁**：区内最大温差超 fZoneDevMax 时锁存 bZoneDevLatch，
 *                              并**强制降零级**（温差失控比缺温更危险）；温差回落到限值 − 迟滞后自动解除。
 *                         串级功率指令（比例段，无积分以免风挡饱和）：
 *                           fCmdPct = Kp · (SP − T_avg) · 级系数，钳 [0, 100]
 *                           级系数：0 级 0.0；1 级 0.4；2 级 0.7；3 级 1.0
 *                         验收向量：
 *                           ① SP=180、四区均 150（Δ=30）且 fDevStage3=20 → 三级，指令 = Kp·30 钳 100
 *                           ② 四区 = {180,181,179,182}（Δ=0）→ 零级，afCmdPct 全 0
 *                           ③ 四区 = {180,180,180,196}（温差 16 > 12）→ 锁存温差联锁 + 强制零级
 *                           ④ 换级后 tStageMin 内偏差剧变 → 级不换（驻留生效）
 * 接口     (Interface)  : 入 bEnable 使能、afTempC 各区实测温度（1..4）、nZoneCnt 有效区数、fSetpointC 设定温度、
 *                         fKpPctPerC 比例增益、fDevStage1/2/3 三级门槛、fZoneDevMaxC 允许最大区间温差、
 *                         fZoneHystC 温差联锁迟滞、tStageMin 最小驻留时长、bReset 复位沿；
 *                         出 afCmdPct 各区加热指令（1..4，钳 0..100）、fAvgTempC 平均温度、
 *                         fZoneDevC 区间最大温差、iStage 当前级（0..3）、bHeating 加热中、
 *                         bZoneDevLatch 温差联锁锁存、eState 相、eCause 成因、bError 故障标志。
 * 边界     (Boundary)   : ① **属主边界（写死）：本件只做"联动分级与温差联锁"，不做单区 PID、
 *                         不驱动固态继电器/调功器**（属单区温控件与 IO 层）；本件输出的是各区统一的
 *                         功率百分比，单区微调由下层温控环叠加；
 *                         ② **分区数组边界**：afTempC / afCmdPct 以字面量上界 4 声明（R104），
 *                         nZoneCnt 作运行时二次闸（钳 1..4），越界区一律输出 0 %；
 *                         ③ **门槛单调闸**：三级门槛须严格递减且为正，温差限与迟滞须为正/非负，违反即锁存 eCfgIllegal；
 *                         ④ **驻留 TON 自复位**：tonDwell 的 IN = 封锁位 ∧ ¬Q（R188），换级即重新封锁；
 *                         ⑤ **温差联锁解除式**：温差 < fZoneDevMaxC − fZoneHystC（自动）∨ bReset 上升沿（人工），
 *                         两式均自证可满足；
 *                         ⑥ 非有限温度样本 → 该区作废（不参与均值与温差），有效区为 0 → 当拍不判、bValid=FALSE；
 *                         ⑦ 零全局耦合、零物理地址。
 * 分工声明 (Scope)      : 本件只管"多温区联动分级与温差联锁"。不接管：单区温度闭环
 *                         （属 FB_DL_DryingOvenZone 族）、层压压力曲线（属 FB_DL_LaminatorPressCtrl）、
 *                         加热器断线诊断（属加热器诊断件）。
 * 来源标签 (Source Tag) : ROADMAP 空勾真缺口 P1（层压机多温区联动，自研 clean-room）
 * 码表     (Codes)      : 本件不占用任何全局数字码位（零码位范式 R297）；诊断由 BOOL + ENUM 出口承担。
 * 红线自检 (Redline)    : R1 ✓ 零 GVL/VAR_EXTERNAL ｜ R2 ✓ 零 %I/%Q/%M ｜ R3 ✓ 纯 IEC 61131-3
 *                         R4 ✓ 分区闸 + 门槛单调闸 + 输出限幅 + 非有限闸 ｜ R5 ✓ 声明逐行同行双语注释
 *                         R6 ✓ ENUM+CASE 含 ELSE 兜底 ｜ R7 ✓ TON/R_TRIG 段 0 无条件刷新
 * 修订历史 (Revision)   : 2026-11-19  v1.0.0  R47 首版（批次 4 · 序号 16）
 *==============================================================================*)

TYPE E_DL_LzsState :
(
    eIdle  := 0,    // 待机相（未使能，指令全 0） / Idle, all commands zero
    eHeat  := 10,   // 升温相（分级投切与温差监视） / Heating, staged switching with deviation supervision
    eFault := 90    // 故障相（组态非法，等复位） / Fault, awaiting reset
);
END_TYPE

TYPE E_DL_LzsCause :
(
    eNone          := 0,   // 无异常 / No anomaly
    eCfgIllegal    := 1,   // 组态非法（区数/门槛/限值越域） / Illegal configuration
    eZoneDevExceed := 2,   // 区间温差超限（锁存，强制零级） / Zone deviation exceeded, latched, forced zero stage
    eSampleBad     := 3,   // 全部区样本非有限（当拍不判） / All zone samples non-finite
    ePhaseBad      := 4    // 非法相位兜底 / Illegal phase fallback
);
END_TYPE

FUNCTION_BLOCK FB_DL_LaminatorZoneSync
VAR_INPUT
    bEnable     : BOOL := FALSE;       // 使能（FALSE 时指令全 0） [-] / Enable, commands zeroed when FALSE
    afTempC     : ARRAY[1..4] OF LREAL;   // 各区实测温度（1..4） [°C] / Zone temperatures, points 1..4
    nZoneCnt    : INT := 4;            // 有效区数，域 1..4 [区] / Active zone count, 1..4
    fSetpointC  : LREAL := 180.0;      // 设定温度 [°C] / Temperature set point [°C]
    fKpPctPerC  : LREAL := 5.0;        // 比例增益，域 > 0 [%/°C] / Proportional gain, > 0
    fDevStage1  : LREAL := 3.0;        // 一级门槛（最小正偏差） [°C] / Stage-1 threshold [°C]
    fDevStage2  : LREAL := 8.0;        // 二级门槛 [°C] / Stage-2 threshold [°C]
    fDevStage3  : LREAL := 20.0;       // 三级门槛（最大） [°C] / Stage-3 threshold [°C]
    fZoneDevMaxC: LREAL := 12.0;       // 允许最大区间温差，域 > 0 [°C] / Maximum allowed inter-zone deviation
    fZoneHystC  : LREAL := 2.0;        // 温差联锁迟滞，域 ≥ 0 [°C] / Deviation latch hysteresis
    tStageMin   : TIME := T#5S;        // 换级最小驻留，域 > T#0S [ms] / Minimum stage dwell time
    bReset      : BOOL := FALSE;       // 故障/锁存复位沿 [-] / Reset edge
END_VAR
VAR_OUTPUT
    afCmdPct    : ARRAY[1..4] OF LREAL;                  // 各区加热指令（钳 0..100） [%] / Zone heater command, 0..100
    fAvgTempC   : LREAL := 0.0;                          // 平均温度（有效区） [°C] / Mean temperature of the valid zones
    fZoneDevC   : LREAL := 0.0;                          // 区间最大温差 [°C] / Maximum inter-zone deviation
    iStage      : INT := 0;                              // 当前投切级（0..3） [级] / Present stage, 0..3
    bHeating    : BOOL := FALSE;                          // 加热中（级 ≥ 1 且未被锁存） [-] / Heating active
    bZoneDevLatch : BOOL := FALSE;                        // 温差联锁锁存 [-] / Deviation interlock, latched
    bValid      : BOOL := FALSE;                          // 判据有效（至少一区有限） [-] / Judgement valid
    eState      : E_DL_LzsState := E_DL_LzsState.eIdle;   // 相出口 [-] / Phase outlet
    eCause      : E_DL_LzsCause := E_DL_LzsCause.eNone;   // 成因出口（R190 归因唯一） [-] / Cause outlet
    bError      : BOOL := FALSE;                          // 故障标志（仅组态级） [-] / Error flag, configuration only
END_VAR
VAR
    _eState   : E_DL_LzsState := E_DL_LzsState.eIdle;    // 内部相（CASE 唯一写入目标） / Internal phase
    _eCause   : E_DL_LzsCause := E_DL_LzsCause.eNone;    // 成因锁存量 / Latched cause
    _bFault   : BOOL := FALSE;                           // 故障锁存位 / Latched fault bit
    _bDevLat  : BOOL := FALSE;                           // 温差联锁锁存位 / Latched deviation bit
    _iStage   : INT := 0;                                // 内部级（驻留保持量） / Internal stage, dwell state
    _bDwellBlk: BOOL := FALSE;                           // 驻留封锁位（换级后置位） / Dwell blocking bit
    _fSum     : LREAL := 0.0;                            // 有效区温度累加 [°C] / Sum of valid zone temperatures
    _fMin     : LREAL := 0.0;                            // 有效区最小温度 [°C] / Minimum valid temperature
    _fMax     : LREAL := 0.0;                            // 有效区最大温度 [°C] / Maximum valid temperature
    _fAvg     : LREAL := 0.0;                            // 平均温度工作值 [°C] / Mean working value
    _fDev     : LREAL := 0.0;                            // 偏差工作值 [°C] / Deviation working value
    _fZoneDev : LREAL := 0.0;                            // 区间温差工作值 [°C] / Inter-zone deviation working value
    _fCmd     : LREAL := 0.0;                            // 指令工作值 [%] / Command working value
    _fStageK  : LREAL := 0.0;                            // 级系数 [-] / Stage gain factor
    _nValid   : INT := 0;                                // 有效区计数 [区] / Valid zone count
    _i        : INT := 0;                                // 区循环下标 / Zone loop index
    _bCfgBad  : BOOL := FALSE;                           // 组态非法当拍量 / Illegal configuration this scan
    _bInit    : BOOL := FALSE;                           // 首区初始化标志（本拍首个有效区） / First-valid-zone flag
    tonDwell  : TON;                                     // 换级驻留实例，段 0 无条件调用 / Stage dwell instance
    rtReset   : R_TRIG;                                  // 复位沿实例，段 0 无条件调用 / Reset edge instance
END_VAR
VAR CONSTANT
    DL_LZS_N      : INT := 4;             // 区数上限（与数组字面量上界同源） [区] / Zone upper bound
    DL_LZS_PCT_MAX: LREAL := 100.0;       // 指令上限 [%] / Command upper bound
    DL_LZS_PCT_MIN: LREAL := 0.0;         // 指令下限 [%] / Command lower bound
    DL_LZS_K1     : LREAL := 0.4;         // 一级级系数 [-] / Stage-1 gain factor
    DL_LZS_K2     : LREAL := 0.7;         // 二级级系数 [-] / Stage-2 gain factor
    DL_LZS_K3     : LREAL := 1.0;         // 三级级系数 [-] / Stage-3 gain factor
    DL_LZS_EPS    : LREAL := 1.0E-9;      // 浮点判等容差 [°C] / Equality tolerance
END_VAR

(* —— 段 0：组态闸 + TON 与沿无条件周期刷新（R228A；驻留 TON 自复位，R188） —— *)
_bCfgBad := (nZoneCnt < 1) OR (nZoneCnt > DL_LZS_N)                                        // 区数须在 1..4 / Zone count within 1..4
         OR (NOT ((fDevStage3 > fDevStage2) AND (fDevStage2 > fDevStage1) AND (fDevStage1 > 0.0)))   // 三级门槛严格递减且为正
         OR (fZoneDevMaxC <= 0.0) OR (fZoneHystC < 0.0) OR (fZoneHystC >= fZoneDevMaxC)     // 温差限与迟滞越域 / Deviation limits
         OR (fKpPctPerC <= 0.0) OR (tStageMin <= T#0S);                                     // 增益与驻留须为正 / Gain and dwell positive
rtReset(CLK := bReset);                                                                     // 复位沿 / Reset edge
tonDwell(IN := _bDwellBlk AND (NOT tonDwell.Q), PT := tStageMin);                            // 换级驻留（自复位振荡） / Stage dwell

(* —— 段 1：单拍/输出量预置（锁存量 _eCause/_bFault/_bDevLat/_iStage/_bDwellBlk 不入清单，R107） —— *)
fAvgTempC     := 0.0;                                                                       // 平均温度预置 / Mean preset
fZoneDevC     := 0.0;                                                                       // 区间温差预置 / Deviation preset
iStage        := 0;                                                                         // 级出口预置 / Stage outlet preset
bHeating      := FALSE;                                                                     // 加热中预置 / Heating preset
bValid        := FALSE;                                                                     // 有效位预置 / Validity preset
bError        := FALSE;                                                                     // 故障标志预清（R45 配对） / Error preset
_fSum := 0.0; _fMin := 0.0; _fMax := 0.0;                                                   // 统计量预置 / Statistics preset
_fAvg := 0.0; _fDev := 0.0; _fZoneDev := 0.0; _fCmd := 0.0; _fStageK := 0.0;                // 工作值预置 / Working values preset
_nValid := 0; _bInit := FALSE;                                                              // 计数与初始化标志预置 / Count and init preset
_i := 1;                                                                                    // 区循环下标归位 / Loop index preset
afCmdPct[1] := DL_LZS_PCT_MIN; afCmdPct[2] := DL_LZS_PCT_MIN;                               // 指令逐区预清零（1/4） / Zone commands preset 1 and 2
afCmdPct[3] := DL_LZS_PCT_MIN; afCmdPct[4] := DL_LZS_PCT_MIN;                               // 指令逐区预清零（3/4） / Zone commands preset 3 and 4

(* —— 段 2：组态闸（非法即锁存） —— *)
IF _bCfgBad THEN
    _eCause := E_DL_LzsCause.eCfgIllegal;                                                   // 归因：组态非法 / Cause: illegal configuration
    _bFault := TRUE;                                                                        // 锁存 / Latch
    _eState := E_DL_LzsState.eFault;                                                        // 入故障相 / Enter fault phase
END_IF

(* —— 段 3：迁出链（bReset 上升沿：清组态故障与温差锁存，R228B） —— *)
IF rtReset.Q THEN
    _bFault  := FALSE;                                                                      // 清故障锁存 / Clear fault latch
    _bDevLat := FALSE;                                                                      // 清温差锁存 / Clear the deviation latch
    _eCause  := E_DL_LzsCause.eNone;                                                        // 清成因 / Clear cause
    _iStage  := 0;                                                                          // 级归零 / Stage cleared
    _eState  := E_DL_LzsState.eIdle;                                                        // 回待机相 / Back to idle
END_IF

(* —— 段 4：相迁移（使能驱动；故障相由段 3 迁出） —— *)
CASE _eState OF

E_DL_LzsState.eIdle:
    IF bEnable AND (NOT _bCfgBad) THEN
        _eState := E_DL_LzsState.eHeat;                                                     // 使能进升温相 / Enter heating
    END_IF

E_DL_LzsState.eHeat:
    IF NOT bEnable THEN
        _iStage := 0;                                                                        // 失能：级归零（指令全 0） / Disable clears the stage
        _eState := E_DL_LzsState.eIdle;                                                     // 回待机相（不借故障相过桥） / Back to idle
    END_IF

E_DL_LzsState.eFault:
    ;                                                                                        // 故障相：由段 3 复位沿迁出 / Exit via the reset edge

ELSE
    _eCause := E_DL_LzsCause.ePhaseBad;                                                      // 归因：非法相位 / Cause: illegal phase
    _bFault := TRUE;                                                                         // 锁存 / Latch
    _eState := E_DL_LzsState.eFault;                                                         // 强拉故障相 / Force fault phase

END_CASE

(* —— 段 5：有效区统计（非有限区作废；区内最大温差） —— *)
IF _eState = E_DL_LzsState.eHeat THEN
    FOR _i := 1 TO DL_LZS_N DO
        IF (_i <= nZoneCnt) AND NOT ((afTempC[_i] <> afTempC[_i]) OR ((afTempC[_i] - afTempC[_i]) <> (afTempC[_i] - afTempC[_i]))) THEN
            _nValid := _nValid + 1;                                                         // 有效区计数 / Valid count
            _fSum := _fSum + afTempC[_i];                                                   // 累加 / Accumulate
            IF (NOT _bInit) OR (afTempC[_i] < _fMin) THEN
                _fMin := afTempC[_i];                                                       // 最小值 / Minimum
            END_IF
            IF (NOT _bInit) OR (afTempC[_i] > _fMax) THEN
                _fMax := afTempC[_i];                                                       // 最大值 / Maximum
            END_IF
            _bInit := TRUE;                                                                 // 首个有效区已处理 / First valid zone handled
        END_IF
    END_FOR

    IF _nValid > 0 THEN
        _fAvg := _fSum / INT_TO_LREAL(_nValid);                                             // 平均（分母已证 ≥ 1） / Mean
        _fZoneDev := _fMax - _fMin;                                                         // 区间温差 / Inter-zone deviation
        _fDev := fSetpointC - _fAvg;                                                        // 偏差（正 = 欠温） / Deviation, positive means below set point
        bValid := TRUE;                                                                     // 判据有效 / Valid

        (* —— 段 6：温差联锁（超限锁存并强制零级；回落过迟滞自动解除） —— *)
        IF (_fZoneDev > fZoneDevMaxC) AND (NOT _bDevLat) THEN
            _bDevLat := TRUE;                                                               // 超限：锁存 / Beyond the limit: latch
            _eCause := E_DL_LzsCause.eZoneDevExceed;                                        // 归因：区间温差超限 / Cause: inter-zone deviation
            _iStage := 0;                                                                   // 强制零级（安全侧优先于升温） / Force stage zero
            _bDwellBlk := TRUE;                                                             // 换级后进入驻留 / Enter dwell
        ELSIF _bDevLat AND (_fZoneDev < (fZoneDevMaxC - fZoneHystC)) THEN
            _bDevLat := FALSE;                                                              // 回落过迟滞：自动解除 / Recovered: auto-release
        END_IF

        (* —— 段 7：分级投切（驻留窗内不换级） —— *)
        IF NOT _bDevLat THEN
            IF (NOT _bDwellBlk) OR tonDwell.Q THEN
                _bDwellBlk := FALSE;                                                        // 驻留窗满：允许换级 / Dwell elapsed
                IF _fDev > fDevStage3 THEN
                    IF _iStage <> 3 THEN
                        _iStage := 3; _bDwellBlk := TRUE;                                    // 升三级并重新驻留 / Stage 3
                    END_IF
                ELSIF _fDev > fDevStage2 THEN
                    IF _iStage <> 2 THEN
                        _iStage := 2; _bDwellBlk := TRUE;                                    // 二级 / Stage 2
                    END_IF
                ELSIF _fDev > fDevStage1 THEN
                    IF _iStage <> 1 THEN
                        _iStage := 1; _bDwellBlk := TRUE;                                    // 一级 / Stage 1
                    END_IF
                ELSE
                    IF _iStage <> 0 THEN
                        _iStage := 0; _bDwellBlk := TRUE;                                    // 零级（保温） / Stage 0
                    END_IF
                END_IF
            END_IF
        END_IF

        (* —— 段 8：串级功率指令（比例段，级系数缩放，逐区钳位） —— *)
        CASE _iStage OF
        1: _fStageK := DL_LZS_K1;                                                            // 一级系数 / Stage-1 factor
        2: _fStageK := DL_LZS_K2;                                                            // 二级系数 / Stage-2 factor
        3: _fStageK := DL_LZS_K3;                                                            // 三级系数 / Stage-3 factor
        ELSE
            _fStageK := 0.0;                                                                 // 零级：无功率 / Stage 0: no power
        END_CASE
        _fCmd := fKpPctPerC * _fDev * _fStageK;                                              // 比例指令 / Proportional command
        IF _fCmd > DL_LZS_PCT_MAX THEN
            _fCmd := DL_LZS_PCT_MAX;                                                         // 上钳 / Clamp high
        ELSIF _fCmd < DL_LZS_PCT_MIN THEN
            _fCmd := DL_LZS_PCT_MIN;                                                         // 下钳（负偏差不制冷） / Clamp low
        END_IF
        IF _bDevLat OR (_iStage = 0) THEN
            _fCmd := DL_LZS_PCT_MIN;                                                         // 锁存或零级：指令归零 / Zero command
        END_IF

        FOR _i := 1 TO DL_LZS_N DO
            IF _i <= nZoneCnt THEN
                afCmdPct[_i] := _fCmd;                                                       // 各区统一指令（联动语义） / Uniform command per zone
            ELSE
                afCmdPct[_i] := DL_LZS_PCT_MIN;                                              // 越界区零指令 / Out-of-range zones zeroed
            END_IF
        END_FOR
    ELSE
        _eCause := E_DL_LzsCause.eSampleBad;                                                  // 归因：全部区非有限（当拍不判） / Cause: all samples invalid
    END_IF
END_IF

(* —— 段 9：出口单点映射（名实双出口，R191） —— *)
fAvgTempC     := _fAvg;                                                                       // 平均温度出口 / Mean outlet
fZoneDevC     := _fZoneDev;                                                                   // 区间温差出口 / Deviation outlet
iStage        := _iStage;                                                                     // 级出口 / Stage outlet
bHeating      := (_iStage >= 1) AND (NOT _bDevLat) AND (_eState = E_DL_LzsState.eHeat);       // 加热中出口 / Heating outlet
bZoneDevLatch := _bDevLat;                                                                    // 温差锁存出口 / Deviation latch outlet
eState        := _eState;                                                                     // 相出口 / Phase outlet
eCause        := _eCause;                                                                     // 成因出口 / Cause outlet
bError        := _bFault;                                                                     // 故障标志 / Error flag

END_FUNCTION_BLOCK

(* ---- FB_DL_LaneDivertCtrl.st ---- *)
(*
    FB_DL_LaneDivertCtrl —— 输送线道岔分流控制器（到件 → 岔口动作 → 尾件确认 → 恢复直行）
    ------------------------------------------------------------------
    组件名称  : FB_DL_LaneDivertCtrl
    分类      : DL_Process / Conveyor
    前缀      : FB_DL_
    版本      : 1.0.0
    溯源      : 借鉴点 —— S-9 输送线工程惯例（R7 先例）的「命令 - 反馈 -
                确认」三段分层骨架，以及 PackML（ISA-TR88.00.02）最小子集
                态命名语义（只借「最小子集 + 明确终止态」的态组织）。
                本件只借**骨架与态组织**，岔口三段判据 / 码位 100% 自有。
                clean-room 声明 —— 零代码行复制；定时与沿检测仅用 IEC 61131-3
                标准库 TON / R_TRIG / F_TRIG。
                许可证 —— 本件 MIT；来源标签 s9-conv 为内部自研线，
                t2-7-packml 仅指公开标准条款，无版权文本继承。
    平台      : 纯 IEC 61131-3，CODESYS 3.5 / TwinCAT 3 / InoProShop / Machine Expert 通用
    作者      : 道莅代码库 · PLC编程专家（R71 构建轮 · 批 2 · 序号 6）
    ------------------------------------------------------------------
    功能说明  : 分流道岔「命令 - 反馈 - 确认」三段顺控：
                eIdle 待机 →（到件上升沿 ∧ 岔口回位 ∧ 分流道空闲）eActuate
                岔口动作（发 bDivertCmd，等 bActDone 反馈）→（bActDone 确认，
                uDivertCount 计数）ePassing 通过（bRelease 放行，等尾件越过 =
                到件信号下降沿，F_TRIG 承载）→ eRestore 回位（撤 bDivertCmd /
                bRelease，等 bActHome）→ eIdle。
                拒放不排队（计划口径）：到件时岔口未回位或分流道占用 →
                拒收计数（信息级 37A4），不缓存到件沿 —— 防积压误分；
                周期内（ePassing）后续到件沿忽略，连续来件最小间隔由到件
                传感器信号本身承载，本件不造额外节拍参数（无魔法数）。
                动作反馈超时归因唯一（R190）：eActuate 等 bActDone 超时 →
                37A1；eRestore 等 bActHome 超时 → 37A2，绝不共用码值；
                超时即故障锁存 + 放行撤销（放行撤销必能在码表找到对应码，
                R45 口径）。
                定时器设计：单实例 _tonPhase，PT 由当前相在段 8 以 IF/ELSIF
                链逐相选择（eActuate / eRestore 两相均用 tActTimeout），**每
                周期无条件调用**（规则 ⑦），相切换时 IN 随条件清零复位，
                **不跨相累计**（定时器纪律：单定时器逐相 PT，已声明选型）。
                起立判据「先判后信」（R42）：eActuate 的 bActDone 为本拍
                复验的实时反馈，不在沿上锁存旧反馈。
    错误码    : 16#0002_37A0 组态非法（tActTimeout 非正，延时不可表示），锁存
                            —— 故障级
                16#0002_37A1 岔口动作反馈超时（eActuate 等 bActDone），锁存 +
                            放行撤销 —— 故障级
                16#0002_37A2 岔口回位反馈超时（eRestore 等 bActHome），锁存
                            —— 故障级
                16#0002_37A3 非法相枚举（CASE ELSE 兜底），锁存 —— 故障级
                16#0002_37A4 到件被拒（岔口未回位或分流道占用），拒放不排队
                            —— 信息级，不置 bError
    码位总账  : 37A0 / 37A1 / 37A2 / 37A3 用（均故障级）
                37A4 用（信息级，bError 恒 FALSE）
    状态机    : ENUM E_DL_LdcPhase 五态，CASE 全覆盖 + ELSE 兜底（锁存 37A3
                回 eFault）。迁移表见功能说明；bReset 上升沿：解锁存 →
                eIdle（唯一可到达的解除边，R188）。
    边界与披露: 一 组态判据：tActTimeout <= T#0S 拦截（TIME 非负语义下的
                   防御性复检，37A0）；布尔输入无非有限面，不设数值闸；
                二 失能 / 故障相输出回夹（R57）：bDivertCmd / bRelease 全清零
                   —— 失能（bEn = FALSE）为操作态不发码、状态回 eIdle、
                   **锁存保留**（R303）；故障相 bError 置位并回放锁存码，
                   两者语义分离；
                三 计数器 uDivertCount / uRejectCount 饱和不回绕（增量前预判，
                   R28-3 口径）；uDivertCount 在 bActDone 确认拍计数（岔口
                   动作完成即视为一次分流成立），uRejectCount 在拒收拍计数；
                四 到件沿 / 尾件沿（R_TRIG / F_TRIG）与复位沿均在段 2 无条件
                   周期刷新（规则 ⑦），不在任何 IF 分支内实例化；
                五 ePassing 中 bRelease 与 bDivertCmd 同拍保持（岔口须保持
                   分流位直至尾件越过），eRestore 首拍即双清零（放行撤销
                   与回位命令同步，不留悬空放行）；
                六 零全局变量、零 VAR_EXTERNAL、零物理地址、零数组下标、无除法。
    分工声明  : FB_DL_PalletZoneMerge（DL_Process，合流汇入）、
                FB_DL_ConveyorJamDetect（DL_Device，堵塞判级诊断）——本件只管
                「分流道岔命令-反馈-确认」三段，不做合流汇入与堵塞判级，
                三者互引分工不互代。
    修订记录  : 2026-11-22 v1.0.0 首次入库（R71 构建轮 · 批 2 · 序号 6）
*)
TYPE E_DL_LdcPhase :
(
    eIdle     := 0,   (* 待机，等下一个到件沿 / idle, waiting for the next arrival edge *)
    eActuate  := 10,  (* 岔口动作相（发分流命令，等到位反馈）/ the actuate phase, the divert command out, waiting for the in-position feedback *)
    ePassing  := 20,  (* 通过相（放行，等尾件越过 = 到件下降沿）/ the passing phase, released, waiting for the tail to pass *)
    eRestore  := 30,  (* 回位相（撤命令，等回位反馈）/ the restore phase, the command withdrawn, waiting for the home feedback *)
    eFault    := 40   (* 故障相（锁存待复位）/ the fault phase, latched for a reset *)
);
END_TYPE

FUNCTION_BLOCK FB_DL_LaneDivertCtrl
VAR_INPUT
    bEn         : BOOL := TRUE;            (* 使能，[标志]，FALSE 时出口清零且状态回待机（R303）/ the enable, FALSE clears the outlets and returns to idle *)
    bReset      : BOOL := FALSE;           (* 故障复位（上升沿有效），[标志] / the fault reset, rising edge effective *)
    bPartArrive : BOOL := FALSE;           (* 到件传感，[标志]，上升沿 = 头件到 / 下沿 = 尾件越过 / the part arrival sensor, rising = head arrived, falling = tail passed *)
    bLaneFree   : BOOL := TRUE;            (* 分流道空闲（上位注入），[标志] / the divert lane free flag, injected by the upper level *)
    bActDone    : BOOL := FALSE;           (* 岔口动作器到位反馈，[标志] / the diverter in-position feedback *)
    bActHome    : BOOL := TRUE;            (* 岔口动作器回位反馈，[标志] / the diverter home feedback *)
    tActTimeout : TIME := T#3S;            (* 动作 / 回位反馈超时，[ms]，须 > T#0S / the actuation and home feedback timeout *)
END_VAR
VAR_OUTPUT
    eState      : E_DL_LdcPhase := E_DL_LdcPhase.eIdle; (* 相状态出口，[相] / the phase outlet *)
    bDivertCmd  : BOOL;                    (* 岔口动作命令，[标志] / the diverter actuation command *)
    bRelease    : BOOL;                    (* 放行，[标志] / the release flag *)
    uDivertCount: UDINT;                   (* 分流完成计数（饱和不回绕）/ the divert counter, saturating *)
    uRejectCount: UDINT;                   (* 到件拒收计数（饱和不回绕）/ the reject counter, saturating *)
    bError      : BOOL;                    (* 故障标志，锁存故障时为 TRUE / the fault flag, raised while latched *)
    nErrCode    : UDINT;                   (* 错误码，0 = 正常，锁存回放 / the error id, 0 = ok, replayed from the latch *)
END_VAR
VAR
    _rtArrive   : R_TRIG;                  (* 到件上升沿实例（无条件调用）/ the arrival rising edge instance *)
    _ftArrive   : F_TRIG;                  (* 尾件越过下降沿实例（无条件调用）/ the tail passed falling edge instance *)
    _rtReset    : R_TRIG;                  (* 复位上升沿实例（无条件调用）/ the reset rising edge instance *)
    _tonPhase   : TON;                     (* 相反馈超时实例（单定时器逐相 PT，无条件调用）/ the phase feedback timeout timer *)
    _ePhase     : E_DL_LdcPhase := E_DL_LdcPhase.eIdle; (* 相状态寄存器 / the internal phase register *)
    _bFault     : BOOL;                    (* 故障锁存位，仅 bReset 上升沿解除 / the latched fault bit *)
    _nCodeLatch : UDINT;                   (* 锁存成因码，故障期回放 / the latched cause code, replayed *)
    _bCfgBad    : BOOL;                    (* 组态非法标志（逐拍重算）/ the configuration fault flag *)
    _bTimerIn   : BOOL;                    (* 相计时器 IN 条件（显式条件）/ the timer IN condition *)
    _tPhasePt   : TIME;                    (* 相计时器 PT 当前值（逐相选择）/ the timer PT for the current phase *)
END_VAR
VAR CONSTANT
    DL_LDC_CMAX : UDINT := 16#FFFF_FFFE;   (* 计数器饱和上限（增量前预判）/ the counter saturation cap, pre-increment check *)
END_VAR

// 段 1｜出口预置（R256 统一出口预置）/ segment 1, preset every outlet
eState       := _ePhase;                   // 相出口先镜像寄存器 / mirror the phase register first
bDivertCmd   := FALSE;                     // 分流命令预清零（活动相内再置位）/ preset the divert command false
bRelease     := FALSE;                     // 放行预清零（通过相内再置位）/ preset the release false
bError       := FALSE;                     // 故障标志预清零 / preset the error flag false
nErrCode     := 0;                         // 错误码预置无错 / preset the code to zero
_bTimerIn    := FALSE;                     // 计时条件预清零 / preset the timer condition false
_tPhasePt    := tActTimeout;               // 计时 PT 预置缺省值 / preset the timer PT to the default

// 段 2｜沿检测实例无条件调用（规则 ⑦）/ segment 2, the edge instances, called unconditionally
_rtArrive(CLK := bPartArrive);             // 到件上升沿，每周期无条件刷新 / the arrival edge, refreshed every scan
_ftArrive(CLK := bPartArrive);             // 尾件下降沿，每周期无条件刷新 / the tail edge, refreshed every scan
_rtReset(CLK := bReset);                   // 复位沿，每周期无条件刷新 / the reset edge, refreshed every scan

// 段 3｜复位解除：唯一可到达的锁存解除边（R188）/ segment 3, the only latch release edge
IF _rtReset.Q THEN                         // 复位上升沿 / the reset rising edge
    _bFault     := FALSE;                  // 解除故障锁存 / release the fault latch
    _nCodeLatch := 0;                      // 清锁存码 / clear the latched code
    _ePhase     := E_DL_LdcPhase.eIdle;    // 回待机相（安全相）/ back to the safe idle phase
END_IF

// 段 4｜组态守卫（边界一）/ segment 4, the configuration guard
_bCfgBad := (tActTimeout <= T#0S);         // 超时非正（TIME 非负语义下的防御复检）/ a non positive timeout

// 段 5｜首次成因锁存（故障期不重推断，回放锁存码，R189）/ segment 5, the first-cause latch
IF NOT _bFault THEN                        // 未锁存才登记成因 / a cause is registered only while not latched
    IF _bCfgBad THEN                       // 组态非法（根因）/ the configuration, the root cause
        _bFault     := TRUE;               // 置锁存 / latch it
        _nCodeLatch := 16#0002_37A0;       // 故障级：组态非法 / fault level: an illegal configuration
        _ePhase     := E_DL_LdcPhase.eFault; // 迁入故障相 / enter the fault phase
    END_IF
END_IF

// 段 6｜相反馈超时 PT 选择与无条件调用（规则 ⑦，选相不依赖可跳过分支）/ segment 6, the timer PT selection and the unconditional call
IF _ePhase = E_DL_LdcPhase.eActuate THEN   // 岔口动作相 / the actuate phase
    _tPhasePt := tActTimeout;              // 到位反馈超时 / the in-position feedback timeout
    _bTimerIn := TRUE;                     // 相内计时有效 / the timer runs
ELSIF _ePhase = E_DL_LdcPhase.eRestore THEN // 回位相 / the restore phase
    _tPhasePt := tActTimeout;              // 回位反馈超时 / the home feedback timeout
    _bTimerIn := TRUE;                     // 相内计时有效 / the timer runs
ELSE                                       // 其余相不参与计时（缺省分支，非状态机 ELSE）/ the other phases do not time
    _tPhasePt := tActTimeout;              // 缺省 PT，保证 PT 恒有定义 / a default PT, always defined
    _bTimerIn := FALSE;                    // 计时条件清零 / the timer condition cleared
END_IF
_tonPhase(IN := _bTimerIn, PT := _tPhasePt); // 每周期无条件调用 / called every scan without exception

// 段 7｜失能相输出回夹（R57 + R303，先于状态机执行）/ segment 7, the disable phase output clamping
IF (NOT bEn) AND (NOT _bFault) THEN        // 失能且无锁存故障（操作态不发码）/ disabled without a latched fault
    _ePhase := E_DL_LdcPhase.eIdle;        // 状态回待机 / back to idle
END_IF                                     // 输出清零由段 1 预置 + 状态机仅在运行许可时执行共同保证

// 段 8｜相状态机（ENUM + CASE + ELSE 兜底，仅运行许可时执行）/ segment 8, the phase machine, run permit only
IF bEn AND NOT _bFault THEN                // 运行许可成立 / the run permit holds
CASE _ePhase OF
    E_DL_LdcPhase.eIdle:                   // 待机相 / the idle phase
        IF _rtArrive.Q THEN                // 到件上升沿 / an arrival rising edge
            IF bActHome AND bLaneFree THEN // 岔口已回位且分流道空闲 / homed and the lane free
                _ePhase := E_DL_LdcPhase.eActuate; // 进入岔口动作相 / enter the actuate phase
            ELSE                           // 未回位或分流道占用 → 拒放不排队 / not homed or occupied, refused, no queue
                IF uRejectCount < DL_LDC_CMAX THEN // 饱和不回绕（增量前预判）/ saturating
                    uRejectCount := uRejectCount + 1; // 拒收计数递增 / increment the reject counter
                END_IF
                nErrCode := 16#0002_37A4;  // 信息级：到件被拒（不置 bError，R45）/ info level: the arrival refused
            END_IF
        END_IF
    E_DL_LdcPhase.eActuate:                // 岔口动作相 / the actuate phase
        bDivertCmd := TRUE;                // 发分流命令 / raise the divert command
        IF bActDone THEN                   // 到位反馈本拍复验成立（R42 先判后信）/ the in-position feedback verified this scan
            IF uDivertCount < DL_LDC_CMAX THEN // 饱和不回绕 / saturating
                uDivertCount := uDivertCount + 1; // 分流计数递增（动作完成即成立）/ increment the divert counter
            END_IF
            _ePhase := E_DL_LdcPhase.ePassing; // 进入通过相 / enter the passing phase
        ELSIF _tonPhase.Q THEN             // 动作反馈超时（归因唯一 37A1）/ the actuation feedback timed out
            _bFault     := TRUE;           // 锁存故障 / latch the fault
            _nCodeLatch := 16#0002_37A1;   // 故障级：动作反馈超时 / fault level: the actuation feedback timed out
            _ePhase     := E_DL_LdcPhase.eFault; // 迁入故障相（命令随预置清零，回夹）/ enter the fault phase
        END_IF
    E_DL_LdcPhase.ePassing:                // 通过相 / the passing phase
        bDivertCmd := TRUE;                // 岔口保持分流位直至尾件越过（边界五）/ hold the diverter until the tail passes
        bRelease   := TRUE;                // 放行 / release
        IF _ftArrive.Q THEN                // 尾件越过（到件信号下降沿承载）/ the tail passed, carried by the falling edge
            _ePhase := E_DL_LdcPhase.eRestore; // 进入回位相 / enter the restore phase
        END_IF                             // 放行撤销在 eRestore 首拍由预置完成（不留悬空放行）
    E_DL_LdcPhase.eRestore:                // 回位相 / the restore phase
        IF bActHome THEN                   // 回位反馈本拍复验成立 / the home feedback verified this scan
            _ePhase := E_DL_LdcPhase.eIdle; // 回待机 / back to idle
        ELSIF _tonPhase.Q THEN             // 回位反馈超时（归因唯一 37A2）/ the home feedback timed out
            _bFault     := TRUE;           // 锁存故障 / latch the fault
            _nCodeLatch := 16#0002_37A2;   // 故障级：回位反馈超时 / fault level: the home feedback timed out
            _ePhase     := E_DL_LdcPhase.eFault; // 迁入故障相 / enter the fault phase
        END_IF
    E_DL_LdcPhase.eFault:                  // 故障相（锁存保持）/ the fault phase, latched
        bError   := TRUE;                  // 故障标志置位 / raise the fault flag
        nErrCode := _nCodeLatch;           // 回放锁存码（不按当下输入重推断）/ replay the latched code
    ELSE                                   // 非法枚举兜底（回安全相 + 置码，规则 ⑥）/ the illegal enumeration guard
        _bFault     := TRUE;               // 置锁存 / latch it
        _nCodeLatch := 16#0002_37A3;       // 故障级：非法相枚举 / fault level: an illegal phase value
        _ePhase     := E_DL_LdcPhase.eFault; // 回安全相（故障相）/ force the safe fault phase
        bError      := TRUE;               // 故障标志置位（禁静默）/ raise the flag
        nErrCode    := _nCodeLatch;        // 回放锁存码 / replay the latched code
END_CASE
END_IF

// 段 9｜出口映射（名实双出口同源，单点写入，R191）/ segment 9, the outlet mapping
eState := _ePhase;                         // 相出口 = 寄存器（段 8 之后不再触碰）/ the phase outlet, not touched after segment 8
IF _bFault THEN                            // 锁存故障相出口补充（含故障入口拍，回夹不留残拍）/ the latched fault supplement, including the entry scan
    bDivertCmd := FALSE;                   // 分流命令清零（回夹执行输出）/ zero the divert command outlet
    bRelease   := FALSE;                   // 放行清零（回夹）/ zero the release outlet
    bError   := TRUE;                      // 故障标志 / the fault flag
    nErrCode := _nCodeLatch;               // 回放锁存码 / replay the latched code
END_IF
END_FUNCTION_BLOCK
